FUNCTION_BLOCK SKILL_Control (* The skill's state machine inside SKILL_Core: what Start, Stop, Abort and Reset do in each state. A client's command reaches it only once SKILL_Gate has accepted it, so here a command is the same from a client or from a parent. Technical: Skill state machine: START, HALT, ABORT, RESET (a client's already decided by SKILL_Gate); Idle 0, Running 1, Stopping 2, Succeeded 3, Failed 4, Aborted 5; RUN starts the execution (CalledByClient: with the Start arguments, else with the parent's values) *)
  (* Standard: 61499-2 *)
  (* Version 0.1, 2026-09-28, Project contributors, AAU Smart Production Lab *)
  PACKAGE modlib;
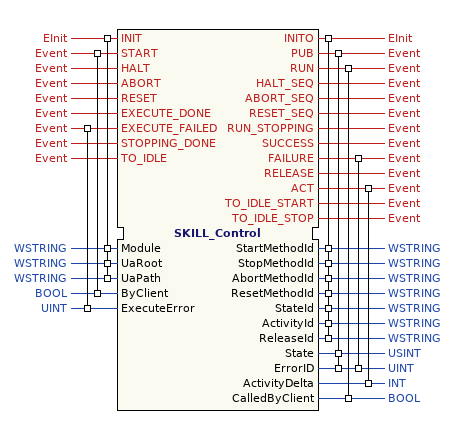
  EVENT_INPUT
    INIT : EInit WITH Module, UaRoot, UaPath; (* Initialise, once at start-up (the INIT chain); takes the values given with it *)
    START WITH ByClient; (* Start a run: a client's Start that SKILL_Gate accepted, or the parent's (ByClient says which) *)
    HALT; (* Stop the run: a client's accepted Stop, or the parent's *)
    ABORT; (* Abort, everything off at once: a client's accepted Abort, or the parent's *)
    RESET; (* Reset from Aborted to Idle: a client's accepted Reset, or the parent's *)
    EXECUTE_DONE; (* The execution ended successfully *)
    EXECUTE_FAILED WITH ExecuteError; (* The execution failed (ExecuteError) *)
    STOPPING_DONE; (* The stop sequence ended *)
    TO_IDLE; (* Succeeded long enough: back to Idle *)
  END_EVENT
  EVENT_OUTPUT
    INITO : EInit WITH StartMethodId, StopMethodId, AbortMethodId, ResetMethodId, StateId, ActivityId, ReleaseId; (* Initialised: the next block of the INIT chain goes on *)
    PUB WITH State, ErrorID; (* Publish State and ErrorID *)
    RUN WITH CalledByClient; (* Run: latch the parameters, start the execution *)
    HALT_SEQ; (* Halt the execute sequence *)
    ABORT_SEQ; (* Abort the sequences *)
    RESET_SEQ; (* Reset the sequences *)
    RUN_STOPPING; (* Run the stop sequence (the skill was stopped) *)
    SUCCESS; (* The run succeeded (the results are set) *)
    FAILURE WITH ErrorID; (* The run failed (ErrorID) *)
    RELEASE; (* A run ended: give up what the skill holds (published if ReleaseAll) *)
    ACT WITH ActivityDelta; (* Count the module's activity (ActivityDelta) *)
    TO_IDLE_START; (* Start the timer back to Idle *)
    TO_IDLE_STOP; (* Stop the timer back to Idle *)
  END_EVENT
  VAR_INPUT
    Module : WSTRING; (* The module's name; its local channels are named after it (loc[<Module>/...]) *)
    UaRoot : WSTRING; (* The module's OPC UA folder, e.g. /Objects/Filling *)
    UaPath : WSTRING; (* This skill's OPC UA folder below UaRoot, e.g. /Skills/Dispensing *)
    ByClient : BOOL; (* The start came from a client over OPC UA (TRUE), or from the parent (FALSE) *)
    ExecuteError : UINT; (* Why the execution failed *)
  END_VAR
  VAR_OUTPUT
    StartMethodId : WSTRING; (* OPC UA ID of the Start method, for its SERVER block *)
    StopMethodId : WSTRING; (* OPC UA ID of the Stop method *)
    AbortMethodId : WSTRING; (* OPC UA ID of the Abort method *)
    ResetMethodId : WSTRING; (* OPC UA ID of the Reset method *)
    StateId : WSTRING; (* OPC UA ID of the published State and ErrorID *)
    ActivityId : WSTRING; (* Local channel of the module's activity count *)
    ReleaseId : WSTRING; (* Local channel the module's equipment is released on *)
    State : USINT; (* Skill state: 0 Idle, 1 Running, 2 Stopping, 3 Succeeded, 4 Failed, 5 Aborted *)
    ErrorID : UINT; (* Error code: 0 none, 1 PreconditionViolated, 2 InvariantViolated, 3 Timeout, 4 NotReady, 5 NotPermitted, 6 Busy, 7 Interrupted, 8 OutOfRange *)
    ActivityDelta : INT; (* +1 when the run starts, -1 when it ends *)
    CalledByClient : BOOL; (* Started over OPC UA (take the Start arguments), not by a parent (take the defaults) *)
  END_VAR
  VAR
    Active : BOOL;
  END_VAR
  EC_STATES
    START;
    Init : Alg_Init -> INITO;
    Idle : Alg_Idle -> PUB;
    Running : Alg_Running -> PUB;
    Stopping : Alg_Stopping -> PUB;
    StopProc : Alg_StopProc -> PUB;
    Succeeded : Alg_Succeeded -> PUB, -> TO_IDLE_START;
    Failed : Alg_Failed -> PUB;
    Aborted : Alg_Aborted -> PUB;
    Go : Alg_Go -> ACT, -> TO_IDLE_STOP, -> RUN;
    Halt : -> HALT_SEQ;
    RunStop : -> RUN_STOPPING;
    Succeed : Alg_Succeed -> ACT, -> RELEASE, -> SUCCESS;
    Fail : Alg_Fail -> ACT, -> RELEASE, -> FAILURE;
    Interrupted : Alg_Interrupted -> ACT, -> RELEASE, -> FAILURE;
    AbortChk;
    AbortActive : Alg_AbortActive -> ABORT_SEQ, -> ACT, -> RELEASE;
    AbortIdle : -> ABORT_SEQ;
    StartRefused : Alg_StartRefused -> FAILURE;
    ResetOk : -> RESET_SEQ;
  END_STATES
  EC_TRANSITIONS
    START TO Init := INIT;
    Init TO Idle := 1;
    Idle TO Go := START;
    Succeeded TO Go := START;
    Failed TO Go := START;
    Aborted TO StartRefused := START;
    StartRefused TO Aborted := 1;
    Running TO Succeed := EXECUTE_DONE;
    Running TO Fail := EXECUTE_FAILED;
    Running TO Halt := HALT;
    Stopping TO RunStop := EXECUTE_DONE;
    Stopping TO RunStop := EXECUTE_FAILED;
    StopProc TO Interrupted := STOPPING_DONE;
    Idle TO AbortChk := ABORT;
    Running TO AbortChk := ABORT;
    Stopping TO AbortChk := ABORT;
    StopProc TO AbortChk := ABORT;
    Succeeded TO AbortChk := ABORT;
    Failed TO AbortChk := ABORT;
    Aborted TO ResetOk := RESET;
    ResetOk TO Idle := 1;
    Go TO Running := 1;
    Halt TO Stopping := 1;
    RunStop TO StopProc := 1;
    Succeed TO Succeeded := 1;
    Succeeded TO Idle := TO_IDLE;
    Fail TO Failed := 1;
    Interrupted TO Failed := 1;
    AbortChk TO AbortActive := [Active];
    AbortChk TO AbortIdle := 1;
    AbortActive TO Aborted := 1;
    AbortIdle TO Aborted := 1;
  END_TRANSITIONS
  ALGORITHM Alg_Init IN ST:
StartMethodId := CONCAT(CONCAT(CONCAT("opc_ua[CREATE_METHOD;", CONCAT(UaRoot, UaPath)), "/Start"), "]");
StopMethodId := CONCAT(CONCAT(CONCAT("opc_ua[CREATE_METHOD;", CONCAT(UaRoot, UaPath)), "/Stop"), "]");
AbortMethodId := CONCAT(CONCAT(CONCAT("opc_ua[CREATE_METHOD;", CONCAT(UaRoot, UaPath)), "/Abort"), "]");
ResetMethodId := CONCAT(CONCAT(CONCAT("opc_ua[CREATE_METHOD;", CONCAT(UaRoot, UaPath)), "/Reset"), "]");
StateId := CONCAT(CONCAT(CONCAT(CONCAT(CONCAT("opc_ua[WRITE;", CONCAT(UaRoot, UaPath)), "/State;"), CONCAT(UaRoot, UaPath)), "/ErrorID"), "]");
ActivityId := CONCAT(CONCAT("loc[", Module), "/activity]");
ReleaseId := CONCAT(CONCAT("loc[", Module), "/release]");
  END_ALGORITHM
  ALGORITHM Alg_Idle IN ST:
State := 0;
  END_ALGORITHM
  ALGORITHM Alg_Running IN ST:
State := 1;
  END_ALGORITHM
  ALGORITHM Alg_Stopping IN ST:
State := 2;
  END_ALGORITHM
  ALGORITHM Alg_StopProc IN ST:
State := 2;
  END_ALGORITHM
  ALGORITHM Alg_Succeeded IN ST:
State := 3;
  END_ALGORITHM
  ALGORITHM Alg_Failed IN ST:
State := 4;
  END_ALGORITHM
  ALGORITHM Alg_Aborted IN ST:
State := 5;
  END_ALGORITHM
  ALGORITHM Alg_Go IN ST:
Active := TRUE;
ActivityDelta := 1;
ErrorID := 0;
CalledByClient := ByClient;
  END_ALGORITHM
  ALGORITHM Alg_Succeed IN ST:
Active := FALSE;
ActivityDelta := -1;
ErrorID := 0;
  END_ALGORITHM
  ALGORITHM Alg_Fail IN ST:
Active := FALSE;
ActivityDelta := -1;
ErrorID := ExecuteError;
  END_ALGORITHM
  ALGORITHM Alg_Interrupted IN ST:
Active := FALSE;
ActivityDelta := -1;
ErrorID := 7;
  END_ALGORITHM
  ALGORITHM Alg_AbortActive IN ST:
Active := FALSE;
ActivityDelta := -1;
ErrorID := 7;
  END_ALGORITHM
  ALGORITHM Alg_StartRefused IN ST:
ErrorID := 4;
  END_ALGORITHM
END_FUNCTION_BLOCK
